FUNCTION_BLOCK TableRotate (* Basic Function Block Type *)
  (* Standard: 61499-2 *)
  (* Version 0.0, 7/2/2026, Template *)
  PACKAGE Main;
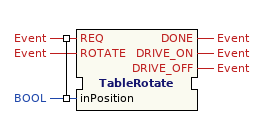
  EVENT_INPUT
    REQ WITH inPosition; (* Normal Execution Request *)
    ROTATE;
  END_EVENT
  EVENT_OUTPUT
    DONE;
    DRIVE_ON;
    DRIVE_OFF;
  END_EVENT
  VAR_INPUT
    inPosition : BOOL; (* Input event qualifier *)
  END_VAR
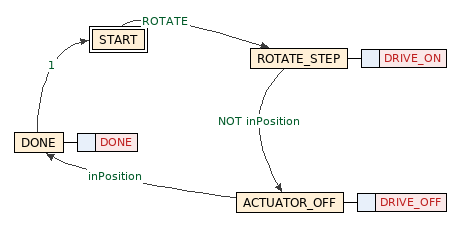
  EC_STATES
    START; (* Initial State *)
    ROTATE_STEP : -> DRIVE_ON;
    ACTUATOR_OFF : -> DRIVE_OFF;
    DONE : -> DONE;
  END_STATES
  EC_TRANSITIONS
    START TO ROTATE_STEP := ROTATE;
    DONE TO START := 1;
    ACTUATOR_OFF TO DONE := inPosition;
    ROTATE_STEP TO ACTUATOR_OFF := NOT inPosition;
  END_TRANSITIONS
  ALGORITHM INIT IN ST: (* Initialization algorithm *)
;
  END_ALGORITHM
  ALGORITHM REQ IN ST: (* Normally executed algorithm *)
;
  END_ALGORITHM
END_FUNCTION_BLOCK
